Fanuc KAREL source: ko00092.KL

-- PROVISIONAL review KL for V770-1; original PC SHA256 f342a6f223502e6bf27e412923b8e36c262440853af8f18a5552b291244e8e4b
-- Incomplete behavior may be omitted. Consult companion uncertainty JSON. Do not deploy.
PROGRAM KO00092
%NOLOCKGROUP
BEGIN
  -- UNRESOLVED_PC offsets 5-12; opcodes 9D,23
  -- UNRESOLVED_PC offsets 17-69; opcodes 27,27,49,7E,AD,27,49,7E,AD,22,31,7E,4A
  -- UNRESOLVED_PC offsets 74-78; opcodes 7F
END KO00092
